TYPE U_APP_CTRL :
UNION
  stCtrl              : ST_TOWER_CTRL;
  byCtrl    AT %Q*    : ARRAY[1..SIZEOF(ST_TOWER_CTRL)] OF BYTE;
END_UNION
END_TYPE

(* stored: Version 1.1.0.1
   DUT U_APP_CTRL: Id {f902224a-8b39-4773-a6df-a85746385b6b} *)
